FUNCTION_BLOCK TestingReset (* CAT Function Block Type *)
  (* Standard: 61499-2 *)
  (* Version 0.0, 11/20/2026, Schneider Electric, template *)
  PACKAGE Main;
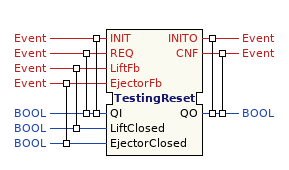
  EVENT_INPUT
    INIT WITH QI; (* Initialization Request *)
    REQ WITH QI; (* Normal Execution Request *)
    LiftFb WITH LiftClosed;
    EjectorFb WITH EjectorClosed;
  END_EVENT
  EVENT_OUTPUT
    INITO WITH QO; (* Initialization Confirm *)
    CNF WITH QO; (* Execution Confirmation *)
  END_EVENT
  VAR_INPUT
    QI : BOOL; (* Input event qualifier *)
    LiftClosed : BOOL;
    EjectorClosed : BOOL;
  END_VAR
  VAR_OUTPUT
    QO : BOOL; (* Output event qualifier *)
  END_VAR
  FBS
    ResetSeq : SeqHead(PermStart := TRUE);
    TR1_TakeOver : SeqStep(TransStepId := 2);
    TR2_AirSlideOff : SeqStep(TransStepId := 3, Exceeded := TRUE);
    TR3_LowerLift : SeqStep(TransStepId := 4);
    TR4_ClearEject : SeqStep(TransStepId := 5);
    TR5_EjectorBack : SeqStep(TransStepId := 6);
    TR_End : SeqTerminate;
    Consts : ANY2ANY_25FC8D56FEEDC9B5(IN1 := TRUE, IN2 := 1, IN3 := 2, IN4 := 0); {SET_ATTRIBUTE(Configuration.GenericFBType.InterfaceParams, Runtime.Standard#CNT:=4;IN${CNT$}:BOOL,INT,INT,INT;OUT${CNT$}:VTQBOOL,VTQINT,VTQINT,VTQINT)}
    OwnerFb : SYMLINKMULTIVARDST_105A0442B8CC61A96(QI := TRUE, NAME1 := 'RES0.Testing.Ejector.sc.progLocal', NAME2 := 'RES0.Testing.AirSlide.sc.progLocal', NAME3 := 'RES0.Testing.Lift.sc.progLocal'); {SET_ATTRIBUTE(Configuration.GenericFBType.InterfaceParams, Runtime.System#I:=3;VALUE${I$}:VTQBOOL,VTQBOOL,VTQBOOL)}
    TakeOverCmd : SYMLINKMULTIVARSRC_105A0442B8CC61A96(QI := TRUE, NAME1 := 'RES0.Testing.Ejector.sc.progLocalSel', NAME2 := 'RES0.Testing.AirSlide.sc.progLocalSel', NAME3 := 'RES0.Testing.Lift.sc.progLocalSel'); {SET_ATTRIBUTE(Configuration.GenericFBType.InterfaceParams, Runtime.System#I:=3;VALUE${I$}:VTQBOOL,VTQBOOL,VTQBOOL)}
    AllLocal : AND_550FE6D62F509EB3(IN3 := TRUE); {SET_ATTRIBUTE(Configuration.GenericFBType.InterfaceParams, Runtime.Standard#CNT:=3;OUT:BOOL)}
    AirSlideOffCmd : SYMLINKMULTIVARSRC_18556BCA74EA878F1(QI := TRUE, NAME1 := 'RES0.Testing.AirSlide.sc.lsp'); {SET_ATTRIBUTE(Configuration.GenericFBType.InterfaceParams, Runtime.System#I:=1;VALUE${I$}:VTQINT)}
    LowerLiftCmd : SYMLINKMULTIVARSRC_18556BCA74EA878F1(QI := TRUE, NAME1 := 'RES0.Testing.Lift.sc.lsp'); {SET_ATTRIBUTE(Configuration.GenericFBType.InterfaceParams, Runtime.System#I:=1;VALUE${I$}:VTQINT)}
    ExtendEjectorCmd : SYMLINKMULTIVARSRC_18556BCA74EA878F1(QI := TRUE, NAME1 := 'RES0.Testing.Ejector.sc.lsp'); {SET_ATTRIBUTE(Configuration.GenericFBType.InterfaceParams, Runtime.System#I:=1;VALUE${I$}:VTQINT)}
    RetractEjectorCmd : SYMLINKMULTIVARSRC_18556BCA74EA878F1(QI := TRUE, NAME1 := 'RES0.Testing.Ejector.sc.lsp'); {SET_ATTRIBUTE(Configuration.GenericFBType.InterfaceParams, Runtime.System#I:=1;VALUE${I$}:VTQINT)}
    EjectTimer : E_DELAY(DT := T#1s);
    EjectLatch : E_SR;
  END_FBS
  EVENT_CONNECTIONS
    INIT TO Consts.REQ;
    Consts.CNF TO ResetSeq.REQ_PERM;
    Consts.CNF TO OwnerFb.INIT;
    Consts.CNF TO TakeOverCmd.INIT;
    Consts.CNF TO AirSlideOffCmd.INIT;
    Consts.CNF TO LowerLiftCmd.INIT;
    Consts.CNF TO ExtendEjectorCmd.INIT;
    Consts.CNF TO RetractEjectorCmd.INIT;
    TR1_TakeOver.STEP_ENTER TO TakeOverCmd.REQ;
    TakeOverCmd.CNF TO AllLocal.REQ;
    OwnerFb.CNF TO AllLocal.REQ;
    AllLocal.CNF TO TR1_TakeOver.TRANS_REQ;
    TR2_AirSlideOff.STEP_ENTER TO AirSlideOffCmd.REQ;
    AirSlideOffCmd.CNF TO TR2_AirSlideOff.TRANS_REQ;
    TR3_LowerLift.STEP_ENTER TO LowerLiftCmd.REQ;
    LowerLiftCmd.CNF TO TR3_LowerLift.TRANS_REQ;
    LiftFb TO TR3_LowerLift.TRANS_REQ;
    TR4_ClearEject.STEP_ENTER TO EjectLatch.R;
    TR4_ClearEject.STEP_ENTER TO ExtendEjectorCmd.REQ;
    ExtendEjectorCmd.CNF TO EjectTimer.START;
    EjectTimer.EO TO EjectLatch.S;
    EjectLatch.EO TO TR4_ClearEject.TRANS_REQ;
    TR4_ClearEject.STEP_LEAVE TO EjectTimer.STOP;
    TR4_ClearEject.STEP_LEAVE TO EjectLatch.R;
    TR5_EjectorBack.STEP_ENTER TO RetractEjectorCmd.REQ;
    RetractEjectorCmd.CNF TO TR5_EjectorBack.TRANS_REQ;
    EjectorFb TO TR5_EjectorBack.TRANS_REQ;
  END_CONNECTIONS
  DATA_CONNECTIONS
    Consts.OUT1 TO TakeOverCmd.VALUE1;
    Consts.OUT1 TO TakeOverCmd.VALUE2;
    Consts.OUT1 TO TakeOverCmd.VALUE3;
    Consts.OUT4 TO AirSlideOffCmd.VALUE1;
    Consts.OUT3 TO LowerLiftCmd.VALUE1;
    Consts.OUT2 TO ExtendEjectorCmd.VALUE1;
    Consts.OUT3 TO RetractEjectorCmd.VALUE1;
    OwnerFb.VALUE1 TO AllLocal.IN1;
    OwnerFb.VALUE2 TO AllLocal.IN2;
    AllLocal.OUT TO TR1_TakeOver.Exceeded;
    LiftClosed TO TR3_LowerLift.Exceeded;
    EjectLatch.Q TO TR4_ClearEject.Exceeded;
    EjectorClosed TO TR5_EjectorBack.Exceeded;
  END_CONNECTIONS
  ADAPTER_CONNECTIONS
    ResetSeq.ISeqChain TO TR1_TakeOver.ISeqChainIn;
    TR1_TakeOver.ISeqChainOut TO TR2_AirSlideOff.ISeqChainIn;
    TR2_AirSlideOff.ISeqChainOut TO TR3_LowerLift.ISeqChainIn;
    TR3_LowerLift.ISeqChainOut TO TR4_ClearEject.ISeqChainIn;
    TR4_ClearEject.ISeqChainOut TO TR5_EjectorBack.ISeqChainIn;
    TR5_EjectorBack.ISeqChainOut TO TR_End.ISeqChainIn;
  END_CONNECTIONS
END_FUNCTION_BLOCK
